// TIA Portal V20 export
// export: Created 2026-10-20T12:45:38.6626938Z, ExportSetting WithDefaults, DisplayName Totally Integrated Automation Portal, DisplayVersion V20 Update 6, DisplayName TIA Portal Openness, DisplayVersion V20 Update 6, DisplayName TIA Portal Version Control Interface, DisplayVersion V20 Update 6, DisplayName SINAMICS Startdrive Advanced, DisplayVersion V20 SP1, DisplayName SINAMICS Startdrive G130, G150, S120, S150, SINAMICS MV, G220, S200, S210, DisplayVersion V20 SP1, DisplayName SINAMICS Startdrive G110M, G120, G120C, G120D, G120P, G115D, DisplayVersion V20 SP1, DisplayName STEP 7 Professional, DisplayVersion V20 Update 6, DisplayName STEP 7 Safety, DisplayVersion V20 Update 2, DisplayName WinCC Basic/Comfort/Advanced, DisplayVersion V20 Update 6, DisplayName WinCC Unified, DisplayVersion V20 Update 6
DATA_BLOCK "OrderTable_HMI_1"   // DB99
{ S7_Optimized_Access := 'TRUE' }
VERSION : 0.1
// stored: AutoNumber true, DBAccessibleFromOPCUA true, IsOnlyStoredInLoadMemory false, IsRetainMemResEnabled false, IsWriteProtectedInAS false, MemoryReserve 100
   VAR
      Start : Bool;
      Pause : Bool;
      Resume : Bool;
      Stop : Bool;
      "Manual order" : Bool;
      Transfer_From_To : Byte;
      "Send VTD Order" : Bool;
      "Send CNV Order" : Bool;
      "Pallet Type" : Byte;
      "Tower 1 Pallet Alignment" : Byte;
      "Tower 2 Pallet Alignment" : Byte;
      "Extractor Pallet Alignment" : Byte;
      "From level" : Byte;
      "To level" : Byte;
      "Testing Time" : UInt;
      "Numer of cycles" : Byte;
      Tower : Byte;
      Level : Byte;
      "Time Running" : UInt;
      Actual_Cycle : Byte;
      "Start Test Visibility" : Bool;
      "Stop Test Visibility" : Bool;
      "Pause Test Visibility" : Bool;
      "Resume Visibility" : Bool;
      "Clear Table Visibility" : Bool;
      "Pallet Type Visibility" : Bool;
      "Tower 1 Visibility" : Bool;
      "Tower 2 Visibility" : Bool;
      "Extractor Visibility" : Bool;
      Auto_Settings_Visibility : Bool;
      "ToExtractor Visibility" : Bool;
      "Manual order Visibility" : Bool;
      "Tower Visibility" : Bool;
      "Level Visibility" : Bool;
      "Send VTD Order Visibility" : Bool;
      "Send CNV Order Visibility" : Bool;
      Clear_OT : Bool;
   END_VAR
BEGIN
END_DATA_BLOCK
